TYPE ST_SpeedControllerStatus :
STRUCT
	velocity 	: LREAL;
	torque		: LREAL;
	homed		: BOOL;
	coupled		: BOOL;
	moving		: BOOL;	
	movingFwd	: BOOL;	
	movingRev	: BOOL;
	faulted		: BOOL;
END_STRUCT
END_TYPE

(* stored: Version 1.1.0.1, ProductVersion 3.1.4024.12
   DUT ST_SpeedControllerStatus: Id {4defb3dd-ea1e-4cfc-b327-55878b6377b9} *)
